(* IEC 61131-3 sources: helmsman/marketing/helmsman-benefits/uploads/mary_had_a_little_lamb, 3 files *)

(* ---- main.st ---- *)
PROGRAM main
VAR_INPUT
  iologik_e1213_di_00 : BOOL;
END_VAR
VAR_OUTPUT
  lamp : BOOL;
  enable : INT;
  slew : DINT;
END_VAR
VAR CONSTANT
  STEPS_PER_REV : DINT := 51200;
  NOTE_SCANS : DINT := 40;
  NOTE_COUNT : DINT := 28;
  NOTE_C : DINT := 40637;
  NOTE_D : DINT := 45619;
  NOTE_G : DINT := 60892;
END_VAR
VAR
  tick : DINT;
  idx : DINT;
END_VAR
  lamp := iologik_e1213_di_00;
  IF iologik_e1213_di_00 THEN
    enable := 1;
    idx := (tick / NOTE_SCANS) MOD NOTE_COUNT;
    tick := tick + 1;
    IF tick >= NOTE_SCANS * NOTE_COUNT THEN
      tick := 0;
    END_IF;
    CASE idx OF
      0: slew := STEPS_PER_REV;
      1: slew := NOTE_D;
      2: slew := NOTE_C;
      3: slew := NOTE_D;
      4: slew := STEPS_PER_REV;
      5: slew := STEPS_PER_REV;
      6: slew := STEPS_PER_REV;
      7: slew := NOTE_D;
      8: slew := NOTE_D;
      9: slew := NOTE_D;
      10: slew := STEPS_PER_REV;
      11: slew := NOTE_G;
      12: slew := NOTE_G;
      13: slew := STEPS_PER_REV;
      14: slew := NOTE_D;
      15: slew := NOTE_C;
      16: slew := NOTE_D;
      17: slew := STEPS_PER_REV;
      18: slew := STEPS_PER_REV;
      19: slew := STEPS_PER_REV;
      20: slew := STEPS_PER_REV;
      21: slew := NOTE_D;
      22: slew := NOTE_D;
      23: slew := STEPS_PER_REV;
      24: slew := NOTE_D;
      25: slew := NOTE_C;
    ELSE
      slew := 0;
    END_CASE;
  ELSE
    tick := 0;
    idx := 0;
    enable := 0;
    slew := 0;
  END_IF;
END_PROGRAM

(* ---- test_lamp_follows_input.st ---- *)
(* lamp turns on when the input goes high and off when it goes low *)
PROGRAM test_lamp_follows_input
VAR_OUTPUT
  iologik_e1213_di_00 : BOOL;
  done : BOOL;
END_VAR
VAR_INPUT
  lamp : BOOL;
END_VAR
VAR
  n : INT;
  lamp_off_first : ASSERT;
  lamp_on : ASSERT;
  lamp_off_after : ASSERT;
END_VAR
  n := n + 1;
  iologik_e1213_di_00 := (n >= 20) AND (n < 60);
  IF n = 10 THEN
    lamp_off_first(COND := NOT lamp);
  END_IF;
  IF n = 40 THEN
    lamp_on(COND := lamp);
  END_IF;
  IF n = 80 THEN
    lamp_off_after(COND := NOT lamp);
    done := TRUE;
  END_IF;
END_PROGRAM

(* ---- test_motor_one_rps.st ---- *)
(* while the input is high the motor is enabled at 1 rev per second (51200 steps/s), and stopped when it drops *)
PROGRAM test_motor_one_rps
VAR_OUTPUT
  iologik_e1213_di_00 : BOOL;
  done : BOOL;
END_VAR
VAR_INPUT
  lamp : BOOL;
  enable : INT;
  slew : DINT;
END_VAR
VAR
  n : INT;
  speed_on : ASSERT;
  enabled_on : ASSERT;
  speed_off : ASSERT;
  enabled_off : ASSERT;
END_VAR
  n := n + 1;
  iologik_e1213_di_00 := (n >= 20) AND (n < 60);
  IF n = 40 THEN
    speed_on(COND := slew = 51200);
    enabled_on(COND := enable = 1);
  END_IF;
  IF n = 80 THEN
    speed_off(COND := slew = 0);
    enabled_off(COND := enable = 0);
    done := TRUE;
  END_IF;
END_PROGRAM
